(* IEC 61131-3 sources: plcassist-cli/packages/volt-lsp-iec/test-corpus/bakon-nano/Device/Plc Logic/Application/Library Manager/L_EtcSlaveConfig, 24 files *)

(* ---- L_ECC_INTERNAL.gvl ---- *)
VAR_GLOBAL
	SMANUFACTURER : STRING := 'Lenze';
	SDEVCLASSINV : STRING := 'Inverter';
END_VAR

(* ---- GETBOOLEANPROPERTY.fun ---- *)
FUNCTION GETBOOLEANPROPERTY : BOOL
VAR_INPUT
	STKEY : WSTRING;
END_VAR
END_FUNCTION

(* ---- GETCOMPANY.fun ---- *)
FUNCTION GETCOMPANY : WSTRING
END_FUNCTION

(* ---- GETNUMBERPROPERTY.fun ---- *)
FUNCTION GETNUMBERPROPERTY : DINT
VAR_INPUT
	STKEY : WSTRING;
END_VAR
END_FUNCTION

(* ---- GETTEXTPROPERTY.fun ---- *)
FUNCTION GETTEXTPROPERTY : WSTRING
VAR_INPUT
	STKEY : WSTRING;
END_VAR
END_FUNCTION

(* ---- GETTEXTPROPERTY2.fun ---- *)
FUNCTION GETTEXTPROPERTY2 : POINTER TO WSTRING
VAR_INPUT
	STKEY : WSTRING;
END_VAR
END_FUNCTION

(* ---- GETTITLE.fun ---- *)
FUNCTION GETTITLE : WSTRING
END_FUNCTION

(* ---- GETVERSION.fun ---- *)
FUNCTION GETVERSION : VERSION
END_FUNCTION

(* ---- GETVERSIONPROPERTY.fun ---- *)
FUNCTION GETVERSIONPROPERTY : VERSION
VAR_INPUT
	STKEY : WSTRING;
END_VAR
END_FUNCTION

(* ---- L_ECC_INITCDFORLENZEINVERTER.fun ---- *)
FUNCTION L_ECC_INITCDFORLENZEINVERTER : BOOL
VAR_INPUT
	PETCSLAVE : POINTER TO ETCSlave;
END_VAR
END_FUNCTION

(* ---- _L_ECC_XXX_DIAGNOSTICS.fb ---- *)
FUNCTION_BLOCK _L_ECC_XXX_DIAGNOSTICS
VAR_INPUT
	XENABLE : BOOL := TRUE;
END_VAR
VAR_OUTPUT
	XBUSY : BOOL;
	XDONE : BOOL;
	XDIAGACTIVE : BOOL;
	XERRORDETECTED : BOOL;
	XERROR : BOOL;
	EERRORID : L_ECC_eError;
END_VAR
VAR
	XBUSY_INT : BOOL := FALSE;
	XDONE_INT : BOOL := FALSE;
	XERROR_INT : BOOL := FALSE;
	EERRORID_INT : L_ECC_eError;
	XDIAGACTIVE_INT : BOOL := FALSE;
	XERRORDETECTED_INT : BOOL := FALSE;
	SCDEVICEINFO_INT : L_ECC_scDeviceInfo;
	PETCSLAVE_INT : POINTER TO L_ETC.ETCSlave;
	PETCSLAVE_MEM : POINTER TO L_ETC.ETCSlave;
	ESTEPPER : _L_ECC_eStepper;
	UIFORLOOP : UINT;
	XINITDONE : BOOL := FALSE;
	ECMASTER : POINTER TO L_IODrvEtherCAT;
	WMASTERSTATE : L_ETC_STATE := L_ETC_STATE.ETC_STATE_NONE;
	FBGETSLAVESTATE : L_ETC_GetSlaveState;
	WSLAVESTATE : L_ETC_STATE := L_ETC_STATE.ETC_STATE_NONE;
	XSDOSTOPONERROR : BOOL := TRUE;
	FBSDOREAD : L_ETC_CoE_SdoRead;
	FBSDOREAD_XEXECUTE_MEM : BOOL;
	ABYSDOREADRAWVALUES : ARRAY [0..uiSdoReadArraySize] OF BYTE;
	SSDOREADPARSEDVALUE : STRING(255);
	DWSDOREADPARSEDVALUE : DWORD;
	FBSDOWRITE : L_ETC_CoE_SdoWrite;
	ABYSDOWRITERAWVALUES : ARRAY [0..uiSdoWriteArraySize] OF BYTE;
	XSDO_READSYSTEMVERSION : BOOL;
	XFIRSTCALL : BOOL := TRUE;
	XREADCOMPONENTINFODONE : BOOL;
	UISDOREADARRAYSIZE : UINT := 127;
	UISDOWRITEARRAYSIZE : UINT := 3;
	UDISDOTIMEOUT : UDINT := 1000;
END_VAR
END_FUNCTION_BLOCK

METHOD GETDEVICECLASS : BOOL
VAR_IN_OUT
	SDEVICECLASS : STRING;
END_VAR
END_METHOD

METHOD INITFIRSTCALL
END_METHOD

METHOD SETCMPINFODATA : BOOL
END_METHOD

METHOD AMAIN
END_METHOD

METHOD ASTATEMACHINE
END_METHOD

METHOD MCHECKDEVICETYPE : BOOL
VAR_INPUT
	DWPRODUCTID : DWORD;
END_VAR
END_METHOD

METHOD MRESETOUTPUTS
END_METHOD

METHOD MSDO_READ : BOOL
VAR_INPUT
	WINDEX : WORD;
	BYSUBINDEX : BYTE;
END_VAR
END_METHOD

METHOD MSDO_WRITE : BOOL
VAR_INPUT
	WINDEX : WORD;
	BYSUBINDEX : BYTE;
	BYSIZE : BYTE;
	DWVALUE : DWORD;
END_VAR
END_METHOD

METHOD MSETETCSLAVE : BOOL
VAR_INPUT
	PETCSLAVE : POINTER TO ETCSlave;
END_VAR
END_METHOD

(* ---- ETCCONFIGPARAXFER.fb ---- *)
FUNCTION_BLOCK ETCCONFIGPARAXFER EXTENDS L_SUDP_UpDownload
VAR_INPUT
	XPREVENTETCOPERATIONALWHENSDOWRITEERROR : BOOL;
END_VAR
VAR
	BYOLDVALUEOFCONTROLINPUT : BYTE := 16#FF;
	WPARAFILESZ : INT;
	INUMBYTESIO : INT;
	IBUFOFFSET : INT;
	BHEADERTEST : BOOL;
	BIOABORTED : BOOL;
	STATE : FILE_STATE := S_INITIALIZE;
	SPARAFILENAME : STRING(255);
	HPARAFILE : CAA.HANDLE;
	ELASTERROR : L_SUDP_ErrorCodes;
	IPARDATASZ : INT;
	IPARRECSZ : INT;
	FGETFS : FILE.GetSize;
	FOPEN : FILE.Open;
	FREAD : FILE.Read;
	FCLOSE : FILE.Close;
	PIOBUFFER : POINTER TO BYTE;
	AYIOBUFFER : ARRAY [0..1000] OF BYTE;
	PPARMREC : POINTER TO L_SUDP_PARM_RECORD;
	PFILEHDR : POINTER TO L_SUDP_PAR_FILE_HDR;
	PPARMDAT : POINTER TO L_SUDP_PAR_DATA_HDR;
	PETCDEV : POINTER TO ETCSlave;
	ECONTROL : L_SUDP_Control;
	PSATTACHEDERRORTXT : POINTER TO STRING;
	SDOWR : L_ETC_CoE_SdoWrite;
	BIGNOREPARAMETER : BOOL;
	BSDOWRITEERROROCCURS : BOOL;
	GETSLAVESTATE : L_ETC_GetSlaveState;
	GETETCMASTERDIAGNOSTIC : L_ETC_GetMasterDiagnostic;
END_VAR
END_FUNCTION_BLOCK

METHOD CLOSEFILE
END_METHOD

METHOD DOWNLOAD
END_METHOD

METHOD IGNOREINDEX : BOOL
VAR_INPUT
	U16INDEX : UINT;
	U16SUBINDEX : UINT;
END_VAR
END_METHOD

METHOD INITIALIZE
VAR_INPUT
	PETCREMDEV : POINTER TO L_ETCSlave;
END_VAR
END_METHOD

METHOD RESETALLSIGNALS
END_METHOD

(* ---- ETCPARAMETERUPLOAD.fb ---- *)
FUNCTION_BLOCK ETCPARAMETERUPLOAD EXTENDS L_SUDP_UpDownload
VAR_INPUT
	DWFILEOFFSETCHECKSUMCALC : DWORD;
END_VAR
VAR
	PETCDEV : POINTER TO ETCSlave;
	ECONTROL : L_SUDP_Control;
	BYOLDVALUEOFCONTROLINPUT : BYTE := 16#FF;
	UPLSTATE : PARAUPLOAD_STATE := PARAUPLOAD_STATE.UPL_INITIALIZE;
	GETSLAVESTATE : L_ETC_GetSlaveState;
	GETETCMASTERDIAGNOSTIC : L_ETC_GetMasterDiagnostic;
	EUPLOADERROR : L_SUDP_ErrorCodes;
	PRMREADWRITEETC : L_SUDP_PRMFile_ReadWrite_ETC;
END_VAR
END_FUNCTION_BLOCK

METHOD INITIALIZE
VAR_INPUT
	PETCREMDEV : POINTER TO L_ETCSlave;
END_VAR
END_METHOD

METHOD PARAUPLOAD
END_METHOD

(* ---- GLOBALTEXTLIST.fb ---- *)
FUNCTION_BLOCK GLOBALTEXTLIST
VAR
	M_TEXTLISTFILE : STRING(255);
	_STNAMESPACE : STRING;
END_VAR
END_FUNCTION_BLOCK

(* ---- L_ECC_CD_DIAGNOSTIC.fb ---- *)
FUNCTION_BLOCK L_ECC_CD_DIAGNOSTIC EXTENDS _L_ECC_XXX_Diagnostics
VAR
	UIACTSLAVECOUNT : UINT := 0;
	UIACTSLAVEINPROGRESS : UINT;
	PSLAVES : ARRAY [1..uicMaxSlaves] OF POINTER TO ETCSlave;
	USISLAVESSTATE : ARRAY [1..uicMaxSlaves] OF USINT;
	XDATAUPDATED : BOOL;
	UICMAXDEPTH : UINT := 10;
	UICMAXSLAVES : UINT := 256;
END_VAR
END_FUNCTION_BLOCK

METHOD ADDSLAVE : BOOL
VAR_INPUT
	PECATSLAVE : POINTER TO ETCSlave;
END_VAR
END_METHOD

METHOD CHECKECATSLAVE : BOOL
VAR_INPUT
	PCHILD : POINTER TO IoConfigConnector;
END_VAR
END_METHOD

METHOD GETDATA : BOOL
VAR_INPUT
	COMPONENTINFOID : UDINT;
	NEXTSTEP : _L_ECC_eStepper;
END_VAR
VAR_IN_OUT
	STEPPER : _L_ECC_eStepper;
END_VAR
END_METHOD

METHOD UPDATECOMPONENTINFO : BOOL
VAR_INPUT
	DATASELECTION : UDINT;
	SDATA : STRING;
END_VAR
END_METHOD

METHOD AMAIN
END_METHOD

METHOD ASTATEMACHINE
END_METHOD

METHOD MCHECKDEVICETYPE : BOOL
VAR_INPUT
	DWPRODUCTID : DWORD;
END_VAR
END_METHOD

(* ---- L_ECC_S131_DIAGNOSTICS.fb ---- *)
FUNCTION_BLOCK L_ECC_S131_DIAGNOSTICS EXTENDS _L_ECC_XXX_Diagnostics
VAR
	SCBUSCOUPLER_INT : L_ECC_scS13x_Coupler;
	ASCIOSLICES_INT : ARRAY [1..uicMaxIOSlices] OF L_ECC_scS13x_IO_Slice;
	XSLICEREGISTERDONCMPDIR : BOOL;
	XSDO_READSLICESERIALNUMBER : BOOL;
	XSDO_READSLICEMXFILE : BOOL;
	WTEXTREFID : WORD;
	WSELECTEDIOSLICE : WORD;
	WRESETIOSLICES : WORD;
	DWERRORREGISTERHARDWARE_INT : DWORD;
	DWERRORREGISTERDIAGNOSTIC_INT : DWORD;
	LWMODULESTATUSDIAGNOSTIC_INT : DWORD;
	DWDISABLEAUTOACK_INT : DWORD;
	DWERRORCODEHARDWARE_INT : DWORD;
	DWERRORCODEDIAGNOSTIC_INT : DWORD;
	BYSLICEERRORSLICE_HARDWARE : BYTE;
	BYSLICEERRORSLICE_DIAGNOSTIC : BYTE;
	XHARDWAREERRORDETECTED_INT : BOOL := FALSE;
	XDIAGNOSTICERRORDETECTED_INT : BOOL := FALSE;
	SPRODUCTVERSION : STRING;
	SSERIALNUMBER : STRING;
	SHWVERSION : STRING;
	SSWVERSION : STRING;
	SMODULEID : STRING;
	UICMAXIOSLICES : UINT := 64;
END_VAR
END_FUNCTION_BLOCK

METHOD GETDEVICECLASS : BOOL
VAR_IN_OUT
	SDEVICECLASS : STRING;
END_VAR
END_METHOD

METHOD INITFIRSTCALL
END_METHOD

METHOD SETSLICECMPINFODATA : BOOL
END_METHOD

METHOD ACYCLICSTATEMACHINE
END_METHOD

METHOD AINITIALIZATIONSTATEMACHINE
END_METHOD

METHOD ASTATEMACHINE
END_METHOD

METHOD MCHECKDEVICETYPE : BOOL
VAR_INPUT
	DWPRODUCTID : DWORD;
END_VAR
END_METHOD

METHOD MCLEARIOSLICEREGISTRATIONS : BOOL
END_METHOD

METHOD MREGISTERIOSLICE : BOOL
VAR_INPUT
	PSCIOSLICE : POINTER TO L_IOSlice;
	BYSLOTNUMBER : BYTE;
END_VAR
END_METHOD

METHOD MRESETOUTPUTS
END_METHOD

METHOD MSETAUTOACKERROR : BOOL
END_METHOD

METHOD MSETDIAGNOSTICERROR : BOOL
VAR_INPUT
	BYSLICE : BYTE := 1;
	ESEVERITY : _L_ECC_eSeverity := _L_ECC_eSeverity.Fault_Log;
	DWERRORID : DWORD := 0;
END_VAR
END_METHOD

(* ---- L_ECC_SAFETY_DIAGNOSTICS.fb ---- *)
FUNCTION_BLOCK L_ECC_SAFETY_DIAGNOSTICS EXTENDS _L_ECC_XXX_Diagnostics
VAR
	SCCPU_1_INT : L_ECC_scC250_CPU;
	SCCPU_2_INT : L_ECC_scC250_CPU;
	XSDO_SLAVEISIOMODULE : BOOL;
	WTEXTREFID : WORD;
	DWERRORREGISTER_INT : DWORD;
	DWSTATEINPUT_MEM : DWORD;
	DWSTATEOUTPUT_MEM : DWORD;
	DWSTATEINPUT_INT : DWORD;
	DWSTATEOUTPUT_INT : DWORD;
	DWERRORCOUNT : DWORD;
	DWCLEARCOUNT : DWORD;
END_VAR
END_FUNCTION_BLOCK

METHOD GETDEVICECLASS : BOOL
VAR_IN_OUT
	SDEVICECLASS : STRING;
END_VAR
END_METHOD

METHOD ASTATEMACHINE
END_METHOD

METHOD MCHECKDEVICETYPE : BOOL
VAR_INPUT
	DWPRODUCTID : DWORD;
END_VAR
END_METHOD

METHOD MDECODESERIALNUMBER : STRING(11)
VAR_INPUT
	DWSERIALNUMBERBITCODED : DWORD;
END_VAR
END_METHOD

METHOD MRESETOUTPUTS
END_METHOD

METHOD MRESETOUTPUTS_ERRORS
END_METHOD

METHOD MSETDIAGNOSTICERROR : BOOL
VAR_INPUT
	ESEVERITY : _L_ECC_eSeverity := _L_ECC_eSeverity.Fault_Log;
	PSCCPUINFO : POINTER TO L_ECC_scC250_CPU;
END_VAR
END_METHOD

(* ---- L_ECC_SCHEDULER.fb ---- *)
FUNCTION_BLOCK L_ECC_SCHEDULER
VAR_INPUT
	XENABLE : BOOL := TRUE;
END_VAR
VAR
	HEVENTUPDATECONFIGURATIONDONE : RTS_IEC_HANDLE;
	HINTERFACEUPDATECONFIGURATIONDONE : RTS_IEC_HANDLE;
	ITFCALLBACK : CmpEventMgr.ICmpEventCallback;
	MYCONNECTOR : POINTER TO IoConfigConnector;
	SCHEDULER : L_ECC_XXX_Diagnostics_Scheduler;
	COMPONENTDIRECTORY : L_ECC_CD_Diagnostic;
	UICMAXDEPTH : UINT := 10;
END_VAR
END_FUNCTION_BLOCK

METHOD CHILDHASDIAGFB : BOOL
VAR_INPUT
	PCHILD : POINTER TO IoConfigConnector;
END_VAR
END_METHOD

METHOD CYCLICCALL : UDINT
END_METHOD

METHOD EVENTCALLBACK : UDINT
VAR_INPUT
	PEVENTPARAM : POINTER TO EventParam;
END_VAR
END_METHOD

METHOD FB_EXIT : BOOL
VAR_INPUT
	BINCOPYCODE : BOOL;
END_VAR
END_METHOD

METHOD FB_INIT : BOOL
VAR_INPUT
	BINITRETAINS : BOOL;
	BINCOPYCODE : BOOL;
END_VAR
END_METHOD

METHOD GETDIAGFBINSTANCE : POINTER TO _L_ECC_XXX_Diagnostics
VAR_INPUT
	PCHILD_ECATSLAVE : POINTER TO IoConfigConnector;
END_VAR
END_METHOD

METHOD GETDIAGSLAVES : BOOL
END_METHOD

METHOD GETDIAGSLAVESRECURSIVE : BOOL
VAR_INPUT
	PFATHER : POINTER TO IoConfigConnector;
	PCONNLIST : POINTER TO IoConfigConnector;
	CONNLISTCOUNT : DINT;
	DWDEPTH : DWORD;
END_VAR
END_METHOD

METHOD GETECATMASTECONNECTOR : BOOL
VAR_IN_OUT
	PECATMASTERCONNECTOR : POINTER TO IoConfigConnector;
END_VAR
END_METHOD

METHOD INITIALIZE : UDINT
VAR_INPUT
	WMODULETYPE : UINT;
	DWINSTANCE : UDINT;
	PCONNECTOR : POINTER TO IoConfigConnector;
END_VAR
END_METHOD

METHOD NODEISECATMASTER : BOOL
VAR_INPUT
	PNODE : POINTER TO IoConfigConnector;
END_VAR
END_METHOD

(* ---- L_ECC_XXX_DIAGNOSTICS_SCHEDULER.fb ---- *)
FUNCTION_BLOCK L_ECC_XXX_DIAGNOSTICS_SCHEDULER
VAR
	ASCHEDULEDATA : ARRAY [1..uicMaxFBs] OF L_ECC_scScheduleData;
	WNUMREGISTEREDFBS : WORD := 0;
	WMAXFBSPERCYCLE_INT : WORD := 1;
	UISCHEDULEIDX : UINT := 1;
	UISCHEDULELOOPCOUNT : UINT := 0;
	UISCHEDULELOOPMAX : UINT := 0;
	ESCHEDULER : _L_ECC_eSchedule := _L_ECC_eSchedule.INIT;
	DWDIAGCYCLECOUNT : DWORD := 0;
	DWDOUBLEREGISTRATIONCOUNT : DWORD := 0;
	UICMAXFBS : UINT := 256;
END_VAR
END_FUNCTION_BLOCK

METHOD AMAIN
END_METHOD

METHOD ASCHEDULE
END_METHOD

METHOD MFBISREGISTERED : BOOL
VAR_INPUT
	PFB_INSTANCE : POINTER TO _L_ECC_XXX_Diagnostics;
END_VAR
END_METHOD

METHOD MINIT : INT
VAR_INPUT
	WMAXFBSPERCYCLE : WORD := 1;
END_VAR
END_METHOD

METHOD MREGISTERFB : BOOL
VAR_INPUT
	PFB_INSTANCE : POINTER TO _L_ECC_XXX_Diagnostics;
END_VAR
END_METHOD

METHOD MSTOPSCHEDULING : BOOL
END_METHOD

(* ---- L_ETCSLAVE.fb ---- *)
FUNCTION_BLOCK L_ETCSLAVE
VAR_OUTPUT
	PETCSLAVE : POINTER TO ETCSlave;
END_VAR
VAR
	ETCSLAVE : ETCSlave;
	M_HLEMACCESS : RTS_IEC_HANDLE;
	PARSETXFER : EtcConfigParaXfer;
	PARSETUPLOAD : EtcParameterUpload;
	ISMANDATORY : BOOL;
	ISPRESENT : BOOL;
	MODULEHANDLER : L_IMHP_IModuleHandler;
END_VAR
END_FUNCTION_BLOCK

METHOD CYCLICCALL : UDINT
END_METHOD

METHOD FB_EXIT : BOOL
VAR_INPUT
	BINCOPYCODE : BOOL;
END_VAR
END_METHOD

METHOD FB_INIT : BOOL
VAR_INPUT
	BINITRETAINS : BOOL;
	BINCOPYCODE : BOOL;
END_VAR
END_METHOD

METHOD INITIALIZE : UDINT
VAR_INPUT
	WMODULETYPE : UINT;
	DWINSTANCE : UDINT;
	PCONNECTOR : POINTER TO IoConfigConnector;
END_VAR
END_METHOD

(* ---- L_ETCSLAVE_S131.fb ---- *)
FUNCTION_BLOCK L_ETCSLAVE_S131 EXTENDS L_ETCSlave
VAR
	HEVENTUPDATECONFIGURATIONDONE : RTS_IEC_HANDLE;
	HINTERFACEUPDATECONFIGURATIONDONE : RTS_IEC_HANDLE;
	ITFCALLBACK : CmpEventMgr.ICmpEventCallback;
	MYCONNECTOR : POINTER TO IoConfigConnector;
	SOWNCOMMPATH : STRING(199);
	WMODULECOUNT : WORD;
	IIOSLICES : ARRAY [1..c_MaxModules] OF POINTER TO L_IOSlice;
	FBS131_DIAGNOSTICS : L_ECC_S131_Diagnostics;
	C_MAXMODULES : WORD := 64;
END_VAR
END_FUNCTION_BLOCK

METHOD CHILDISIOSLICE : BOOL
VAR_INPUT
	PCHILD : POINTER TO IoConfigConnector;
END_VAR
END_METHOD

METHOD CYCLICCALL : UDINT
END_METHOD

METHOD EVENTCALLBACK : UDINT
VAR_INPUT
	PEVENTPARAM : POINTER TO EventParam;
END_VAR
END_METHOD

METHOD FB_EXIT : BOOL
VAR_INPUT
	BINCOPYCODE : BOOL;
END_VAR
END_METHOD

METHOD FB_INIT : BOOL
VAR_INPUT
	BINITRETAINS : BOOL;
	BINCOPYCODE : BOOL;
END_VAR
END_METHOD

METHOD GETIOSLICEINSTANCE : POINTER TO L_IOSlice
VAR_INPUT
	PCHILD_IOSLICE : POINTER TO IoConfigConnector;
END_VAR
END_METHOD

METHOD GETIOSLICES : BOOL
END_METHOD

METHOD INITIALIZE : UDINT
VAR_INPUT
	WMODULETYPE : UINT;
	DWINSTANCE : UDINT;
	PCONNECTOR : POINTER TO IoConfigConnector;
END_VAR
END_METHOD

METHOD READOWNCOMMPATH : BOOL
END_METHOD

METHOD REGISTERIOSLICE : BOOL
VAR_INPUT
	PSCIOSLICE : POINTER TO L_IOSlice;
	BYSLOTNUMBER : BYTE;
END_VAR
END_METHOD

METHOD WRITEDIAGINSTANCEADDRESS : BOOL
VAR_INPUT
	PCONNECTOR : POINTER TO IoConfigConnector;
END_VAR
END_METHOD

(* ---- L_ETCSLAVE_SAFETY.fb ---- *)
FUNCTION_BLOCK L_ETCSLAVE_SAFETY EXTENDS ETCSlave
VAR_OUTPUT
	PETCSLAVE : POINTER TO ETCSlave;
END_VAR
VAR
	ETCSLAVE : REFERENCE TO ETCSlave;
	FBSAFETYDIAGNOSTICS : L_ECC_Safety_Diagnostics;
END_VAR
END_FUNCTION_BLOCK

METHOD FB_EXIT : BOOL
VAR_INPUT
	BINCOPYCODE : BOOL;
END_VAR
END_METHOD

METHOD FB_INIT : BOOL
VAR_INPUT
	BINITRETAINS : BOOL;
	BINCOPYCODE : BOOL;
END_VAR
END_METHOD

METHOD INITIALIZE : UDINT
VAR_INPUT
	WMODULETYPE : UINT;
	DWINSTANCE : UDINT;
	PCONNECTOR : POINTER TO IoConfigConnector;
END_VAR
END_METHOD

METHOD WRITEDIAGINSTANCEADDRESS : BOOL
VAR_INPUT
	PCONNECTOR : POINTER TO IoConfigConnector;
END_VAR
END_METHOD

METHOD FB_REINIT : BOOL
END_METHOD

(* ---- L_IOSLICE.fb ---- *)
FUNCTION_BLOCK L_IOSLICE
VAR
	MODULEHANDLERBASE : L_IMHP_ModuleHandler := STRUCT(CompActiveDefault := TRUE, Layer := L_IMHP_Layer.Communication, CompType := L_IMHP_ComponentType.EtherCATSlave, DefaultRelationship := L_IMHP_RelationshipID.CommunicationView);
	MODULEID : L_ECC_eDeviceType;
	UIACTUALERROR : UINT;
	REGISTERONCOMPONENTDIRECTORY : L_IC1P_RegisterOnComponentDirectory;
	MYWMODULETYPE : UINT;
	MYDWINSTANCE : UDINT;
	MYPCONNECTOR : POINTER TO IoConfigConnector;
	MODULEHANDLER : L_IMHP_IModuleHandler;
END_VAR
END_FUNCTION_BLOCK

METHOD FB_INIT : BOOL
VAR_INPUT
	BINITRETAINS : BOOL;
	BINCOPYCODE : BOOL;
END_VAR
END_METHOD

METHOD INITIALIZE : UDINT
VAR_INPUT
	WMODULETYPE : UINT;
	DWINSTANCE : UDINT;
	PCONNECTOR : POINTER TO IoConfigConnector;
END_VAR
END_METHOD

METHOD READMODULEID : BOOL
VAR_INPUT
	PCONNECTOR : POINTER TO IoConfigConnector;
END_VAR
END_METHOD

METHOD WRITEINSTANCEADDRESS : BOOL
VAR_INPUT
	PCONNECTOR : POINTER TO IoConfigConnector;
END_VAR
END_METHOD

METHOD MDIAGNOSTICERRORTOERRORCODE : UINT
VAR_INPUT
	EDEVICETYPE : L_ECC_eDeviceType;
	DWERRORID : DWORD := 0;
END_VAR
END_METHOD

METHOD MERRORHANDLER : BOOL
VAR_INPUT
	ESEVERITY : _L_ECC_eSeverity := _L_ECC_eSeverity.Fault_Log;
	DWERRORID : DWORD := 0;
	WTEXTREFID : WORD;
END_VAR
END_METHOD

METHOD MSETCOMMPATH : BOOL
VAR_INPUT
	SPATH : STRING(199);
END_VAR
END_METHOD

(* ---- L_SUDP_PRMFILE_READWRITE_ETC.fb ---- *)
FUNCTION_BLOCK L_SUDP_PRMFILE_READWRITE_ETC EXTENDS L_SUDP_PRMFile_ReadWrite
VAR
	SDORD : L_ETC_CoE_SdoRead;
	FILESIZECHANGED : BOOL;
END_VAR
END_FUNCTION_BLOCK

METHOD BEFORESTARTEXECUTION
END_METHOD

METHOD READVALUEFROMFIELDBUS_LOOP : INT
END_METHOD

METHOD READVALUEFROMFIELDBUS_START
VAR_INPUT
	PARAMHDR : POINTER TO L_SUDP.L_SUDP_PARM_HDR;
	PBYBUFFER : POINTER TO BYTE;
	SZBUFFERSIZE : UINT;
END_VAR
END_METHOD
